FUNCTION_BLOCK JanelaIntertravamento (* Janela de intertravamento: TRUE com o intertravamento ativo e ate TempoDepois apos ele sair *)
  (* Standard: 61499-2 *)
  (* Version 1.1, 05/11/2026, Hidryco, Hidryco, 1.1: eventos de saida listados no ECAction (sem isso o runtime nao emite nenhum; o ST so liga/desliga). 1.0: Janela = intertravamento ativo OU contando TempoDepois (10 s) depois que ele sai. Usado no Motor_VS para o intertravamento nao deixar o equipamento pedindo reset. *)
  PACKAGE SE.Nereda;
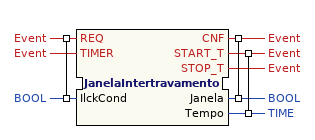
  EVENT_INPUT
    REQ WITH IlckCond; (* Intertravamento mudou *)
    TIMER; (* Fim do tempo (E_DELAY.EO) *)
  END_EVENT
  EVENT_OUTPUT
    CNF WITH Janela; (* Janela mudou *)
    START_T WITH Tempo; (* Inicia o tempo (E_DELAY.START) *)
    STOP_T; (* Cancela o tempo (E_DELAY.STOP) *)
  END_EVENT
  VAR_INPUT
    IlckCond : BOOL; (* Intertravamento ativo *)
  END_VAR
  VAR_OUTPUT
    Janela : BOOL; (* Intertravamento ativo ou recem-saido *)
    Tempo : TIME; (* Tempo do E_DELAY *)
  END_VAR
  VAR
    contando : BOOL; (* Contando o tempo depois do intertravamento *)
    TempoDepois : TIME := T#10s; (* Quanto tempo a janela continua depois que o intertravamento sai *)
  END_VAR
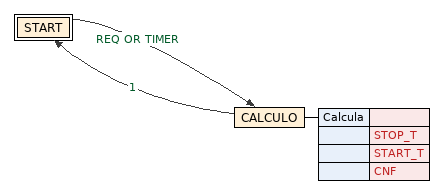
  EC_STATES
    START; (* Estado inicial *)
    CALCULO : Calcula, -> STOP_T, -> START_T, -> CNF; (* Calcula; o algoritmo decide quais eventos saem *)
  END_STATES
  EC_TRANSITIONS
    START TO CALCULO := REQ OR TIMER;
    CALCULO TO START := 1;
  END_TRANSITIONS
  ALGORITHM Calcula IN ST: (* Janela de intertravamento: TRUE com o intertravamento ativo e ate TempoDepois apos ele sair *)
CNF := FALSE;
START_T := FALSE;
STOP_T := FALSE;
IF REQ THEN
    IF IlckCond THEN
        IF contando THEN
            STOP_T := TRUE;
            contando := FALSE;
        END_IF;
        IF NOT Janela THEN
            Janela := TRUE;
            CNF := TRUE;
        END_IF;
    ELSIF Janela AND NOT contando THEN
        (* saiu do intertravamento: segura a janela por TempoDepois *)
        contando := TRUE;
        Tempo := TempoDepois;
        START_T := TRUE;
    END_IF;
ELSIF TIMER THEN
    IF contando THEN
        contando := FALSE;
        IF NOT IlckCond THEN
            Janela := FALSE;
            CNF := TRUE;
        END_IF;
    END_IF;
END_IF;
  END_ALGORITHM
END_FUNCTION_BLOCK
